Fanuc KAREL source: compact_preamble.KL

PROGRAM KB00010
%NOLOCKGROUP
VAR
P1 : STRING[80];P2 : STRING[80];P3:INTEGER;P4:INTEGER;P5 : STRING[80];P6:INTEGER
BEGIN
P1='A'
P2='A'
P3=1
P4=1
P5='A'
P6=1
ATT_WINDOW_D(P1,P2,P3,P4,P5,P6)
END KB00010
